(* IEC 61131-3 sources: Codesys_IAP/Demo/PLC1/Magazijn Overzetter Simulatie Structured Text 2V1_tekst/Programma Structured Text/Structures, 4 files *)

(* ---- hmiIO.st ---- *)
(*#### DECLARATIE ####*)
// Datum : 17 december 2020, Auteur: Gerard Harkema
TYPE hmiIO :
STRUCT
	// Indrukken resetknop
	Ix_Resetknop			: REFERENCE TO BOOL;
	// Keuzeknop staat op hand
	Ix_Hand					: REFERENCE TO BOOL;
	// Keuzeknop staat op auto
	Ix_Auto					: REFERENCE TO BOOL;
	// Indrukken noodstop
	Ix_Noodstop				: REFERENCE TO BOOL;
	// Bekers magazijn zijn op

	// Indrukken startknop
	Ix_Stopknop				: REFERENCE TO BOOL;
	// Indrukken stopknop
	Ix_Startknop			: REFERENCE TO BOOL;
	//Perslucht is aanwezig

	// Visualisatie invisible Gele vlak
	Qx_GeleLamp				: REFERENCE TO BOOL;
	// Visualisatie invisible groene vlak
	Qx_GroeneLamp			: REFERENCE TO BOOL;
	// Visualisatie invisible rode vlak
	Qx_RodeLamp				: REFERENCE TO BOOL;

END_STRUCT
END_TYPE

(* ---- magazijnIO.st ---- *)
(*#### DECLARATIE ####*)
// Datum : 17 december 2020, Auteur: Gerard Harkema
TYPE magazijnIO :
STRUCT
	// Bekers magazijn zijn op
	Ix_MagazijnLeeg				: REFERENCE TO BOOL;
	// Beker is uit dekselmagazijn gestoten
	Ix_UitstoterBekerIn			: REFERENCE TO BOOL;
	// Uitstoter Beker haalt nieuwe beker op
	Ix_UitstoterBekerUit		: REFERENCE TO BOOL;
	// Beker uit magazijn stoten
	Qx_BekerUitstoten			: REFERENCE TO BOOL;

	//Perslucht is aanwezig
	Ix_PersluchtAanwezig 		: REFERENCE TO BOOL;

END_STRUCT
END_TYPE

(* ---- overzetterIO.st ---- *)
(*#### DECLARATIE ####*)
// Datum : 17 december 2020, Auteur: Gerard Harkema
TYPE overzetterIO :
STRUCT
	//Werkstuk door overzetter opgepakt
	Ix_VacuumAanwezig 		:REFERENCE TO BOOL;
	//Overzetter haalt beker op(linker pos.)
	Ix_OverzetterIsLinks 	:REFERENCE TO BOOL;
	//Overzetter plaatst beker op sorteerpositie
	Ix_OverzetterIsRechts 	:REFERENCE TO BOOL;
	//Beker aanwezig op detectiepositie

		//Beker oppakken
	Qx_VacuumAan 			:REFERENCE TO BOOL;
	//Beker loslaten
	Qx_BekerLossen 			:REFERENCE TO BOOL;
	//Overzetter naar bekermagazijn
	Qx_OverzetterLinks 		:REFERENCE TO BOOL;
	//Overzetter naar sorteerpositie
	Qx_OverzetterRechts 	:REFERENCE TO BOOL;

END_STRUCT
END_TYPE

(* ---- stationIO.st ---- *)
(*#### DECLARATIE ####*)
// Datum : 26 november 2026, Auteur: Gerard Harkema
TYPE stationIO :
STRUCT
	// IO van het magazijn
	magazijn		: magazijnIO;
	// IO van de overzetter
	overzetter		: overzetterIO;
END_STRUCT
END_TYPE
